Fanuc KAREL source: KT00595.KL

PROGRAM KT00595
%NOLOCKGROUP
VAR
  R1: REAL
  S2: STRING[80]
  OUT: STRING[80]
BEGIN
  R1 = 2.0
    S2 = 'B'
  OUT = R1 + S2
END KT00595
